Yaskawa INFORM job: ---JEFFRESS-S-SHAPE.JBI

/JOB
//NAME ---JEFFRESS-S-SHAPE
///FOLDERNAME FOLDER052
//POS
///NPOS 8,0,0,0,0,0
///TOOL 0
///POSTYPE PULSE
///PULSE
C00000=28401,16455,-73182,127097,-29642,-144792
C00001=28401,16455,-73182,127097,-29642,-144792
C00002=37465,22609,-75368,139978,-33219,-162115
C00003=8001,27161,-71504,152088,-19686,-162620
C00004=28964,12568,-88664,152226,-29379,-171485
C00005=53108,44,-100427,143060,-40152,-172300
C00006=16689,-3565,-104432,163336,-24118,-177806
C00007=-27964,-12691,-100843,122667,-2858,-119110
//INST
///DATE 2024/07/23 17:24
///ATTR SC,RW
///GROUP1 RB1
NOP
MOVL C00000 V=7.8
MOVL C00001 V=25.0
MOVC C00002 V=25.0
MOVC C00003 V=25.0
MOVC C00004 V=25.0 FPT
MOVC C00005 V=25.0
MOVC C00006 V=25.0
MOVL C00007 V=7.8
END
